// SIMATIC S7-200 project (STEP 7-Micro/WIN), CPU 226 CN REL 02.01

SYMBOL_TABLE USUARIO1
boton1           I1.3
boton2           I1.2
selector         I1.5
act1             Q0.0
act2             Q0.4
act3             Q0.5
act4             Q0.6
END_SYMBOL_TABLE

ORGANIZATION_BLOCK Bloque_de_programa:OB1
TITLE=COMENTARIOS DEL PROGRAMA
BEGIN
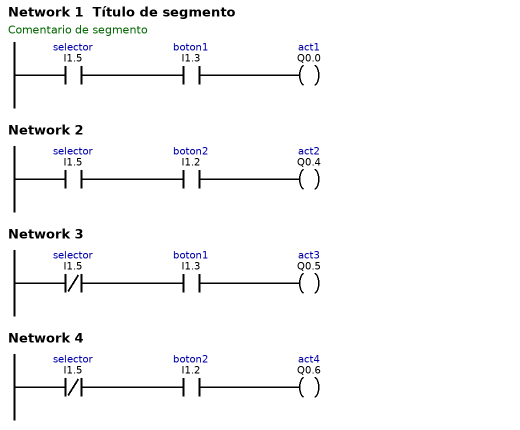
Network 1 // Título de segmento
// Comentario de segmento
// (network saved uncompiled; LAD cells follow)
// row 0: c0 -| |- selector:I1.5  c1 -| |- boton1:I1.3  c2 -( ) act1:Q0.0
Network 2
// (network saved uncompiled; LAD cells follow)
// row 0: c0 -| |- selector:I1.5  c1 -| |- boton2:I1.2  c2 -( ) act2:Q0.4
Network 3
// (network saved uncompiled; LAD cells follow)
// row 0: c0 -|/|- selector:I1.5  c1 -| |- boton1:I1.3  c2 -( ) act3:Q0.5
Network 4
// (network saved uncompiled; LAD cells follow)
// row 0: c0 -|/|- selector:I1.5  c1 -| |- boton2:I1.2  c2 -( ) act4:Q0.6
END_ORGANIZATION_BLOCK
